(* IEC 61131-3 sources: plc-st-coding-agent/agent_dev_r9_stage3/datasets/selfmade/tests, 15 files *)

(* ---- self-easy-01.reference.st ---- *)
FUNCTION_BLOCK FB
VAR_INPUT
    enable : BOOL;
    values : ARRAY[1..8] OF INT;
    count : INT;
    avgEnable : BOOL;
END_VAR
VAR_OUTPUT
    avgOut : REAL;
END_VAR
VAR
    i : INT;
    n : INT;
    sum : DINT;
    keep : REAL;
END_VAR

(* 先把有效样本数裁剪到 [0, 8]，负数和超长都收敛到合法范围 *)
n := count;
IF n < 0 THEN
    n := 0;
ELSIF n > 8 THEN
    n := 8;
END_IF

(* 要点：输出变量在每周期扫描开头就被赋成本周期的计算结果，
   "保持不变"没法靠"不写它"实现——必须先读回旧值再决定写不写。
   这里用静态变量 keep 记住上一周期的有效结果。 *)
IF enable AND avgEnable AND n > 0 THEN
    sum := 0;
    FOR i := 1 TO n DO
        sum := sum + values[i];
    END_FOR
    keep := DINT_TO_REAL(sum) / INT_TO_REAL(n);
END_IF
avgOut := keep;
END_FUNCTION_BLOCK

(* ---- self-easy-02.reference.st ---- *)
FUNCTION_BLOCK FB
VAR_INPUT
    tankLevel : REAL;
    outletFlow : REAL;
    inletPermit : BOOL;
    resetBtn : BOOL;
END_VAR
VAR_OUTPUT
    pumpRun : BOOL;
    alarmHigh : BOOL;
    alarmLow : BOOL;
    outletValveOpen : BOOL;
END_VAR
VAR
    resetEdgeInputPrev : BOOL;
    resetEdge : BOOL;
    latchReset : BOOL;
END_VAR

(* 复位只取上升沿：按住不放只生效一次 *)
resetEdge := resetBtn AND NOT resetEdgeInputPrev;
resetEdgeInputPrev := resetBtn;
latchReset := resetEdge;

(* 报警自保持：置位优先于复位，且复位条件只在上升沿成立一个周期 *)
IF tankLevel >= 85.0 AND NOT latchReset THEN
    alarmHigh := TRUE;
END_IF
IF latchReset THEN
    alarmHigh := FALSE;
END_IF
IF tankLevel <= 15.0 AND NOT latchReset THEN
    alarmLow := TRUE;
END_IF
IF latchReset THEN
    alarmLow := FALSE;
END_IF

(* 联锁：任一报警存在都不得进料 *)
pumpRun := inletPermit AND NOT alarmHigh AND NOT alarmLow
           AND tankLevel < 85.0 AND tankLevel >= 15.0;

(* 出口阀在低液位报警时强制关闭 *)
outletValveOpen := NOT alarmLow AND tankLevel > 15.0;
END_FUNCTION_BLOCK

(* ---- self-hard-01.reference.st ---- *)
FUNCTION_BLOCK FB
VAR_INPUT
    flowLow : BOOL;
    ackBtn : BOOL;
    sensorOK : BOOL;
END_VAR
VAR_OUTPUT
    alarmActive : BOOL;
    alarmAcked : BOOL;
    highHigh : BOOL;
END_VAR
VAR
    ackEdgeInputPrev : BOOL;
    ackEdge : BOOL;
    alarmState : INT;
END_VAR

ackEdge := ackBtn AND NOT ackEdgeInputPrev;
ackEdgeInputPrev := ackBtn;

(* 高优先级：传感器断线，独立判定，不被低优先级抑制 *)
highHigh := NOT sensorOK;

(* 0 正常；1 激活未确认；2 激活已确认；3 条件消失但仍待人工确认。
   题面第2条把状态3的 alarmAcked 也定义为 TRUE。 *)
CASE alarmState OF
    0:
        IF flowLow THEN alarmState := 1; END_IF
    1:
        IF NOT flowLow THEN alarmState := 3; END_IF
    2:
        IF NOT flowLow THEN alarmState := 0; END_IF
    3:
        IF flowLow THEN alarmState := 1; END_IF
END_CASE
IF ackEdge THEN
    IF flowLow THEN
        alarmState := 2;
    ELSE
        alarmState := 0;
    END_IF
END_IF
alarmActive := alarmState <> 0;
alarmAcked := (alarmState = 2) OR (alarmState = 3);
END_FUNCTION_BLOCK

(* ---- self-hard-02.reference.st ---- *)
FUNCTION_BLOCK FB
VAR_INPUT
    startBtn : BOOL;
    abortBtn : BOOL;
    setpoint : REAL;
    pv : REAL;
    maxDuration : INT;
END_VAR
VAR_OUTPUT
    elapsed : INT;
    phase : INT;
    timeout : BOOL;
END_VAR
VAR
    startEdgeInputPrev : BOOL;
    startEdge : BOOL;
END_VAR

(* phase: 0=空闲 1=升温 2=保温 9=中止/超时结束 *)
startEdge := startBtn AND NOT startEdgeInputPrev;
startEdgeInputPrev := startBtn;

IF startEdge THEN
    phase := 1;
    elapsed := 0;
    timeout := FALSE;
ELSIF abortBtn THEN
    phase := 9;
ELSIF phase = 1 OR phase = 2 THEN
    (* 计时靠扫描周期自累加，不依赖外部时钟 *)
    elapsed := elapsed + 1;
    (* 阶段推进：升温到设定值转保温；已是保温则保持 *)
    IF phase = 1 AND pv >= setpoint THEN
        phase := 2;
    END_IF
    (* 超时判定放在阶段推进之后，保证"到设定值"的优先级低于"超时停机" *)
    IF elapsed >= maxDuration THEN
        timeout := TRUE;
        phase := 9;
    END_IF
END_IF
END_FUNCTION_BLOCK

(* ---- self-hard-03.reference.st ---- *)
FUNCTION_BLOCK FB
VAR_INPUT
    pushEn : BOOL;
    pushItem : INT;
    popEn : BOOL;
END_VAR
(* fifo 由调用方分配、FB 内部读写，必须是 VAR_IN_OUT；写成 VAR_INPUT 就成了
   只读形参，往里面写会被静态检查直接拒掉（E_WRITE_INPUT）。 *)
VAR_IN_OUT
    fifo : ARRAY[1..8] OF INT;
END_VAR
VAR_OUTPUT
    count : INT;
    full : BOOL;
    empty : BOOL;
    head : INT;
END_VAR
VAR
    pushPrev : BOOL;
    popPrev : BOOL;
    pushEdge : BOOL;
    popEdge : BOOL;
    wr : INT := 1;
    rd : INT := 1;
END_VAR

(* 边沿 = 本周期电平 且 上次周期不是这个电平。
   把"上次电平"和"本周期边沿"分两个变量存，别把边沿算回同一个变量：
   pushEdge := pushEn AND NOT pushEdge 这种写法把边沿覆盖掉上次电平，
   一旦电平连续两个周期为真（如 q7 同周期出队+入队），第二周期算不出边沿，
   入队被静默丢弃。 *)
pushEdge := pushEn AND NOT pushPrev;
popEdge := popEn AND NOT popPrev;
pushPrev := pushEn;
popPrev := popEn;

(* 出队：空队列忽略。先把"这一笔算数"的判断用局部变量兜住，
   因为下面 count := count - 1 已经改变了判断依据。 *)
IF popEdge AND count > 0 THEN
    count := count - 1;
    rd := rd + 1;
    IF rd > 8 THEN
        rd := 1;
    END_IF
END_IF

(* 入队：满队列丢弃。入队判定用**出队之后**的 count，
   所以同一周期既有出队又有入队时，这一格是真的能腾出来用的。 *)
IF pushEdge AND count < 8 THEN
    fifo[wr] := pushItem;
    count := count + 1;
    wr := wr + 1;
    IF wr > 8 THEN
        wr := 1;
    END_IF
END_IF

(* 队列空了指针才归位。必须放在出入队之后，而且要精确到"本周期结束时
   真正空了"；写在这个位置、用 count = 0 判定即可：上面的入队已经执行完，
   同一周期出队腾空又入队时 count 不会是 0，不会被误清零。 *)
IF count <= 0 THEN
    rd := 1;
    wr := 1;
END_IF

full := count >= 8;
empty := count <= 0;
IF empty THEN
    head := 0;
ELSE
    head := fifo[rd];
END_IF
END_FUNCTION_BLOCK

(* ---- self-hard-04.reference.st ---- *)
FUNCTION_BLOCK FB
VAR_INPUT
    demand : INT;
    runHours : ARRAY[1..5] OF LINT;
    rotated : BOOL;
END_VAR
VAR_OUTPUT
    leadPump : INT;
    lagPump : INT;
    runningCount : INT;
END_VAR
VAR
    i : INT;
    j : INT;
    need : INT;
    tmp : LINT;
    order : ARRAY[1..5] OF INT;
END_VAR

(* 需求先裁剪到 0..5，否则后面按 order[i] 取泵号会越界 *)
need := demand;
IF need < 0 THEN
    need := 0;
ELSIF need > 5 THEN
    need := 5;
END_IF

(* 选择排序：按运行小时升序得到泵号次序 *)
FOR i := 1 TO 5 DO
    order[i] := i;
END_FOR
FOR i := 1 TO 4 DO
    FOR j := i + 1 TO 5 DO
        IF runHours[order[j]] < runHours[order[i]] THEN
            tmp := order[i];
            order[i] := order[j];
            order[j] := tmp;
        END_IF
    END_FOR
END_FOR

runningCount := need;
IF need = 0 THEN
    leadPump := 0;
    lagPump := 0;
ELSIF need = 1 THEN
    leadPump := order[1];
    lagPump := 0;
ELSE
    leadPump := order[1];
    lagPump := order[2];
    (* 均衡轮换：两台泵小时数差小于阈值 50 时互换主备，
       让备泵有机会顶上去，避免主泵长期独挑磨损。 *)
    IF rotated AND (runHours[order[2]] - runHours[order[1]]) < 50 THEN
        leadPump := order[2];
        lagPump := order[1];
    END_IF
END_IF
END_FUNCTION_BLOCK

(* ---- self-hard-05.reference.st ---- *)
FUNCTION_BLOCK FB
VAR_INPUT
 runRequest : BOOL;
 flameOK : BOOL;
 o2Valid : BOOL;
 o2PV : REAL;
 baseAir : REAL;
 resetBtn : BOOL;
END_VAR
VAR_OUTPUT
 fuelPermit : BOOL;
 trimEnable : BOOL;
 airTrim : REAL;
 airCommand : REAL;
 tripLatched : BOOL;
 o2Fault : BOOL;
END_VAR
VAR
 prevReset : BOOL;
 tripMem : BOOL;
END_VAR
o2Fault := (NOT o2Valid) OR (o2PV < 0.0) OR (o2PV > 21.0);
IF runRequest AND NOT flameOK THEN
 tripMem := TRUE;
ELSIF resetBtn AND NOT prevReset AND NOT runRequest AND NOT flameOK THEN
 tripMem := FALSE;
END_IF;
prevReset := resetBtn;
tripLatched := tripMem;
fuelPermit := runRequest AND flameOK AND NOT tripMem;
trimEnable := fuelPermit AND NOT o2Fault;
IF trimEnable THEN
 airTrim := 2.0 * (2.0 - o2PV);
 IF airTrim > 10.0 THEN airTrim := 10.0; END_IF;
 IF airTrim < -10.0 THEN airTrim := -10.0; END_IF;
ELSE
 airTrim := 0.0;
END_IF;
IF fuelPermit THEN
 airCommand := baseAir + airTrim;
 IF airCommand > 100.0 THEN airCommand := 100.0; END_IF;
 IF airCommand < 0.0 THEN airCommand := 0.0; END_IF;
ELSE
 airCommand := 0.0;
END_IF;
END_FUNCTION_BLOCK

(* ---- self-hard-06.reference.st ---- *)
FUNCTION_BLOCK FB
VAR_INPUT
 runRequest : BOOL;
 pressure : REAL;
 pressureValid : BOOL;
 fuelFlow : REAL;
 steamFlow : REAL;
 outletCmd : INT;
 outletFeedback : INT;
 resetBtn : BOOL;
END_VAR
VAR_OUTPUT
 tripLatched : BOOL;
 fuelPermit : BOOL;
 currentCauseMask : WORD;
 latchedCauseMask : WORD;
 diagnosticActive : BOOL;
END_VAR
VAR
 prevReset : BOOL;
 tripMem : BOOL;
 latMem : WORD;
 valveCnt : INT;
END_VAR
currentCauseMask := 0;
IF resetBtn AND NOT prevReset AND NOT runRequest AND pressureValid
 AND (pressure <= 4200.0) THEN
 tripMem := FALSE;
 latMem := 0;
 valveCnt := 0;
END_IF;
prevReset := resetBtn;
IF NOT runRequest THEN
 valveCnt := 0;
ELSIF NOT pressureValid THEN
 currentCauseMask := 16#0001;
 valveCnt := 0;
 tripMem := TRUE;
ELSIF pressureValid AND (pressure >= 4500.0) THEN
 IF (outletCmd >= 50) AND (outletFeedback <= 10) THEN
  valveCnt := valveCnt + 1;
  IF valveCnt > 3 THEN valveCnt := 3; END_IF;
 ELSE
  valveCnt := 0;
 END_IF;
 IF valveCnt >= 3 THEN
  currentCauseMask := currentCauseMask OR 16#0002;
 END_IF;
 IF (fuelFlow >= 4.0) AND (steamFlow <= 10.0) THEN
  currentCauseMask := currentCauseMask OR 16#0004;
 END_IF;
 IF currentCauseMask = 0 THEN
  currentCauseMask := 16#0008;
 END_IF;
 tripMem := TRUE;
ELSE
 valveCnt := 0;
END_IF;
IF tripMem THEN
 latMem := latMem OR currentCauseMask;
END_IF;
tripLatched := tripMem;
latchedCauseMask := latMem;
diagnosticActive := (currentCauseMask <> 0);
fuelPermit := runRequest AND NOT tripMem;
END_FUNCTION_BLOCK

(* ---- self-hard-07.reference.st ---- *)
FUNCTION_BLOCK FB
VAR_INPUT
 mode : INT;
 resetBtn : BOOL;
 dt : REAL;
 tempSP : REAL;
 tempPV : REAL;
 flowPV : REAL;
 manualFlowSP : REAL;
 manualValve : REAL;
END_VAR
VAR_OUTPUT
 flowSP : REAL;
 valveCommand : REAL;
 fault : BOOL;
 normalMode : BOOL;
END_VAR
VAR
 prevReset : BOOL;
 initDone : BOOL;
 lastMode : INT;
 accT : REAL;
 accF : REAL;
 oFlow : REAL;
 oValve : REAL;
 eTemp : REAL;
 eFlow : REAL;
 trial : REAL;
 normalMem : BOOL;
END_VAR
fault := (mode < 0) OR (mode > 2) OR (dt <= 0.0) OR (dt > 10.0);
normalMem := FALSE;
IF (NOT initDone) OR (resetBtn AND NOT prevReset) OR fault THEN
 oFlow := manualFlowSP;
 oValve := manualValve;
 accT := oFlow - 1.0 * (tempSP - tempPV);
 accF := oValve - 2.0 * (oFlow - flowPV);
 lastMode := mode;
 initDone := TRUE;
ELSIF lastMode <> mode THEN
 IF mode <> 2 THEN
  oFlow := manualFlowSP;
 END_IF;
 accT := oFlow - 1.0 * (tempSP - tempPV);
 accF := oValve - 2.0 * (oFlow - flowPV);
 lastMode := mode;
ELSE
 normalMem := TRUE;
 IF mode = 0 THEN
  oFlow := manualFlowSP;
  oValve := manualValve;
  accT := oFlow - 1.0 * (tempSP - tempPV);
  accF := oValve - 2.0 * (oFlow - flowPV);
 ELSIF mode = 1 THEN
  oFlow := manualFlowSP;
  accT := oFlow - 1.0 * (tempSP - tempPV);
  eFlow := oFlow - flowPV;
  trial := accF + 0.5 * eFlow * dt;
  oValve := 2.0 * eFlow + trial;
  IF oValve > 100.0 THEN oValve := 100.0; END_IF;
  IF oValve < 0.0 THEN oValve := 0.0; END_IF;
  accF := oValve - 2.0 * eFlow;
 ELSE
  eTemp := tempSP - tempPV;
  trial := accT + 0.2 * eTemp * dt;
  oFlow := 1.0 * eTemp + trial;
  IF oFlow > 50.0 THEN oFlow := 50.0; END_IF;
  IF oFlow < 0.0 THEN oFlow := 0.0; END_IF;
  accT := oFlow - 1.0 * eTemp;
  eFlow := oFlow - flowPV;
  trial := accF + 0.5 * eFlow * dt;
  oValve := 2.0 * eFlow + trial;
  IF oValve > 100.0 THEN oValve := 100.0; END_IF;
  IF oValve < 0.0 THEN oValve := 0.0; END_IF;
  accF := oValve - 2.0 * eFlow;
 END_IF;
END_IF;
prevReset := resetBtn;
flowSP := oFlow;
valveCommand := oValve;
normalMode := normalMem;
END_FUNCTION_BLOCK

(* ---- self-medium-01.reference.st ---- *)
(* 配方结构体必须显式定义：题目给的是 ARRAY[1..8] OF ST_Recipe，
   没有 TYPE 块就读不到字段名，结构体成员访问会被直接判错。 *)
TYPE ST_Recipe :
STRUCT
    recipeID : INT;
    totalRatio : REAL;
    temperature : REAL;
END_STRUCT
END_TYPE

FUNCTION_BLOCK FB
VAR_INPUT
    recipe : ARRAY[1..8] OF ST_Recipe;
    selSlot : INT;
    loadCmd : BOOL;
    running : BOOL;
END_VAR
VAR_OUTPUT
    valid : BOOL;
    loadedID : INT;
END_VAR
VAR
    loadEdgeInputPrev : BOOL;
    loadEdge : BOOL;
    ok : BOOL;
    slotOK : BOOL;
    r : ST_Recipe;
END_VAR

loadEdge := loadCmd AND NOT loadEdgeInputPrev;
loadEdgeInputPrev := loadCmd;
(* 生产运行中不接受装载命令：连有效位都不刷新，保持上一次判定 *)
IF loadEdge AND NOT running THEN
    slotOK := (selSlot >= 1) AND (selSlot <= 8);
    (* 关键：先判槽位合法再访问数组。IEC 的 AND 不保证短路，
       所以不能写成 "slotOK AND recipe[selSlot].xxx" 这种依赖短路的写法 *)
    valid := FALSE;
    IF slotOK THEN
        r := recipe[selSlot];
        ok := r.recipeID <> 0;
        IF r.totalRatio < 99.0 OR r.totalRatio > 101.0 THEN
            ok := FALSE;
        END_IF
        IF r.temperature < 30.0 OR r.temperature > 180.0 THEN
            ok := FALSE;
        END_IF
        valid := ok;
        IF ok THEN
            loadedID := r.recipeID;
        END_IF
    END_IF
END_IF
END_FUNCTION_BLOCK

(* ---- self-medium-02.reference.st ---- *)
FUNCTION_BLOCK FB
VAR_INPUT
    enable : BOOL;
    rawValue : REAL;
END_VAR
VAR_OUTPUT
    filteredValue : REAL;
    windowFull : BOOL;
    sampleCount : INT;
END_VAR
VAR
    buf : ARRAY[1..8] OF REAL;
    wr : INT;
    i : INT;
    sum : REAL;
    keep : REAL;
END_VAR

(* 关断时清空历史，但输出保持最后一次的有效值 *)
IF NOT enable THEN
    FOR i := 1 TO 8 DO
        buf[i] := 0.0;
    END_FOR
    wr := 0;
    sampleCount := 0;
    windowFull := FALSE;
ELSE
    (* 环形缓冲：wr 指向最老元素，写进去就等于淘汰最老的那个 *)
    wr := wr + 1;
    IF wr > 8 THEN
        wr := 1;
    END_IF
    buf[wr] := rawValue;
    IF sampleCount < 8 THEN
        sampleCount := sampleCount + 1;
    END_IF
    windowFull := sampleCount >= 8;

    (* 只对**实际已有**的样本求平均，未满时不得按 0 填充 *)
    sum := 0.0;
    FOR i := 1 TO sampleCount DO
        sum := sum + buf[i];
    END_FOR
    keep := sum / INT_TO_REAL(sampleCount);
END_IF
(* 每一拍都从静态变量刷新输出：输出变量本身不记忆，靠 keep 记忆 *)
filteredValue := keep;
END_FUNCTION_BLOCK

(* ---- self-medium-03.reference.st ---- *)
FUNCTION_BLOCK FB
VAR_INPUT
    openBtn : BOOL;
    closeBtn : BOOL;
    openLimit : BOOL;
    closeLimit : BOOL;
    obstacle : BOOL;
END_VAR
VAR_OUTPUT
    motorUp : BOOL;
    motorDown : BOOL;
    errorFlag : BOOL;
END_VAR
VAR
    state : INT;
    openPrev : BOOL;
    closePrev : BOOL;
    openEdge : BOOL;
    closeEdge : BOOL;
END_VAR

(* 状态编码：0=IDLE 1=OPENING 2=CLOSING 3=FAULT *)
openEdge := openBtn AND NOT openPrev;
openPrev := openBtn;
closeEdge := closeBtn AND NOT closePrev;
closePrev := closeBtn;

(* 障碍优先于一切：无论哪个方向，立即停机 *)
IF obstacle THEN
    motorUp := FALSE;
    motorDown := FALSE;
    IF state <> 3 THEN
        IF state = 2 THEN
            state := 1;
        ELSE
            state := 3;
            errorFlag := TRUE;
        END_IF
    END_IF
ELSE
    (* 障碍解除后必须能重新启动：FAULT 只是"停着等"，不是永久锁死。
       这一段必须写在 ELSE 里——写进 IF obstacle 里面就成了"只有还挡着
       的时候才放行"，语义完全反了。
       但**不能在这里清 errorFlag**：清锁存和"允许动作"必须是同一件事，
       否则会出现"errorFlag 还亮着电机已经转起来"的中间状态，
       直接违反 S4（G(errorFlag -> !motorUp & !motorDown)）。
       所以锁存只在真正接受指令、状态从 IDLE 迁出时清除。 *)
    CASE state OF
        0:
            IF openEdge AND NOT openLimit THEN
                state := 1;
                errorFlag := FALSE;
            ELSIF closeEdge AND NOT closeLimit THEN
                state := 2;
                errorFlag := FALSE;
            END_IF
        1:
            IF openLimit THEN
                state := 0;
            END_IF
        2:
            IF closeLimit THEN
                state := 0;
            END_IF
        3:
            (* 故障锁存：按第 8 条，只有两键同按才算人工复位。
               障碍消失只是"可以复位了"，不是"已经复位"——
               否则障碍消失的那一拍就会允许起机，违反第 7 条。 *)
            IF openBtn AND closeBtn THEN
                state := 0;
                errorFlag := FALSE;
            END_IF
    END_CASE

    (* 电机输出由状态唯一决定，互锁保证不会同时两个方向 *)
    motorUp := (state = 1);
    motorDown := (state = 2);
END_IF
END_FUNCTION_BLOCK

(* ---- self-medium-04.reference.st ---- *)
FUNCTION_BLOCK FB
VAR_INPUT
    startBtn : BOOL;
    resetBtn : BOOL;
    doneSensor : BOOL;
    targetVol : REAL;
    flowVol : REAL;
END_VAR
VAR_OUTPUT
    valveOpen : BOOL;
    fillsToday : INT;
END_VAR
VAR
    resetEdgeInputPrev : BOOL;
    startEdgeInputPrev : BOOL;
    startEdge : BOOL;
    resetEdge : BOOL;
    accumulated : REAL;
    filling : BOOL;
    waitAck : BOOL;
END_VAR

startEdge := startBtn AND NOT startEdgeInputPrev;
startEdgeInputPrev := startBtn;
resetEdge := resetBtn AND NOT resetEdgeInputPrev;
resetEdgeInputPrev := resetBtn;

(* 复位最高优先级：清零计数、关阀 *)
IF resetEdge THEN
    fillsToday := 0;
    valveOpen := FALSE;
    filling := FALSE;
    waitAck := FALSE;
    accumulated := 0.0;
ELSE
    (* 运途中重复按启动无效：只在非灌装、非待确认时接受 *)
    (* 待确认期间再按启动：允许直接开灌下一瓶，上一瓶未确认就不计数了 *)
    IF startEdge AND waitAck THEN
        waitAck := FALSE;
    END_IF
    IF startEdge AND NOT filling THEN
        filling := TRUE;
        valveOpen := TRUE;
        accumulated := 0.0;
    END_IF

    IF filling THEN
        accumulated := accumulated + flowVol;
        (* 达到或超过目标立即关阀，用 >= 而不是 > *)
        IF accumulated >= targetVol THEN
            valveOpen := FALSE;
            filling := FALSE;
            waitAck := TRUE;
        END_IF
    END_IF

    (* 计数只在满瓶确认之后发生一次 *)
    IF waitAck AND doneSensor THEN
        fillsToday := fillsToday + 1;
        waitAck := FALSE;
    END_IF
END_IF
END_FUNCTION_BLOCK

(* ---- self-medium-05.reference.st ---- *)
FUNCTION_BLOCK FB
VAR_INPUT
 enable : BOOL;
 resetBtn : BOOL;
 dt : LREAL;
 steamFlow : LREAL;
 fuelFlow : LREAL;
 steamTemp : LREAL;
 steamPressure : LREAL;
END_VAR
VAR_OUTPUT
 qualified : BOOL;
 dataFault : BOOL;
 qualifiedTon : LREAL;
 fuelTon : LREAL;
 revenue : LREAL;
 cost : LREAL;
 netProfit : LREAL;
END_VAR
VAR
 prevReset : BOOL;
 qTon : LREAL;
 fTon : LREAL;
END_VAR
qualified := (steamTemp >= 447.0) AND (steamTemp <= 453.0)
 AND (steamPressure >= 3750.0) AND (steamPressure <= 3850.0);
dataFault := (dt <= 0.0) OR (dt > 10.0)
 OR (steamFlow < 0.0) OR (steamFlow > 90.0)
 OR (fuelFlow < 0.0) OR (fuelFlow > 6.0);
IF resetBtn AND NOT prevReset THEN
 qTon := 0.0;
 fTon := 0.0;
ELSIF enable AND NOT dataFault THEN
 fTon := fTon + fuelFlow * dt / 1000.0;
 IF qualified THEN
  qTon := qTon + steamFlow * dt / 1000.0;
 END_IF;
END_IF;
prevReset := resetBtn;
qualifiedTon := qTon;
fuelTon := fTon;
revenue := qTon * 280.0;
cost := fTon * 1500.0;
netProfit := revenue - cost;
END_FUNCTION_BLOCK

(* ---- self-medium-06.reference.st ---- *)
FUNCTION_BLOCK FB
VAR_INPUT
 enable : BOOL;
 resetBtn : BOOL;
 sensorValid : BOOL;
 setpoint : REAL;
 temperature : REAL;
 dt : REAL;
 bias : REAL;
END_VAR
VAR_OUTPUT
 power : REAL;
 correction : REAL;
 fault : BOOL;
END_VAR
VAR
 prevReset : BOOL;
 prevE : REAL;
 hasHist : BOOL;
 eNow : REAL;
 eDe : REAL;
 xx : REAL;
 yy : REAL;
 mx : REAL;
 zx : REAL;
 px : REAL;
 my : REAL;
 zy : REAL;
 py : REAL;
 wsum : REAL;
 wc : REAL;
 cOut : REAL;
 edgeReset : BOOL;
END_VAR
fault := (NOT sensorValid) OR (dt <= 0.0) OR (dt > 10.0);
edgeReset := resetBtn AND NOT prevReset;
IF edgeReset OR (NOT enable) OR fault THEN
 cOut := 0.0;
 hasHist := FALSE;
 prevE := 0.0;
ELSE
 eNow := setpoint - temperature;
 IF hasHist THEN
  eDe := (eNow - prevE) / dt;
 ELSE
  eDe := 0.0;
 END_IF;
 xx := eNow / 10.0;
 IF xx > 1.0 THEN xx := 1.0; END_IF;
 IF xx < -1.0 THEN xx := -1.0; END_IF;
 yy := eDe / 2.0;
 IF yy > 1.0 THEN yy := 1.0; END_IF;
 IF yy < -1.0 THEN yy := -1.0; END_IF;
 mx := MAX(-xx, 0.0);
 zx := 1.0 - ABS(xx);
 px := MAX(xx, 0.0);
 my := MAX(-yy, 0.0);
 zy := 1.0 - ABS(yy);
 py := MAX(yy, 0.0);
 wsum := mx * my + mx * zy + mx * py + zx * my + zx * zy + zx * py
  + px * my + px * zy + px * py;
 wc := mx * my * (-30.0) + mx * zy * (-20.0) + mx * py * (-10.0)
  + zx * my * (-10.0) + zx * zy * 0.0 + zx * py * 10.0
  + px * my * 10.0 + px * zy * 20.0 + px * py * 30.0;
 IF wsum > 0.0 THEN
  cOut := wc / wsum;
 ELSE
  cOut := 0.0;
 END_IF;
 prevE := eNow;
 hasHist := TRUE;
END_IF;
prevReset := resetBtn;
correction := cOut;
IF edgeReset OR (NOT enable) OR fault THEN
 power := 0.0;
ELSE
 power := bias + cOut;
 IF power > 100.0 THEN power := 100.0; END_IF;
 IF power < 0.0 THEN power := 0.0; END_IF;
END_IF;
END_FUNCTION_BLOCK
